// TIA Portal V20 export
// export: Created 2026-10-20T18:54:16.3544517Z, ExportSetting None, DisplayName Totally Integrated Automation Portal, DisplayVersion V20 Update 6, DisplayName TIA Portal Openness, DisplayVersion V20 Update 6, DisplayName TIA Portal Version Control Interface, DisplayVersion V20 Update 6, DisplayName SINAMICS Startdrive Advanced, DisplayVersion V20 SP1, DisplayName SINAMICS Startdrive G130, G150, S120, S150, SINAMICS MV, G220, S200, S210, DisplayVersion V20 SP1, DisplayName SINAMICS Startdrive G110M, G120, G120C, G120D, G120P, G115D, DisplayVersion V20 SP1, DisplayName STEP 7 Professional, DisplayVersion V20 Update 6, DisplayName STEP 7 Safety, DisplayVersion V20 Update 2, DisplayName WinCC Basic/Comfort/Advanced, DisplayVersion V20 Update 6, DisplayName WinCC Unified, DisplayVersion V20 Update 6
VAR_GLOBAL   // PLC tag table "IO_Main Panel"
   "MAIN PANEL STACK LIGHT RED" AT %Q350.0 : Bool;   // TESTED
   "MAIN PANEL STACK LIGHT AMBER" AT %Q350.1 : Bool;   // TESTED
   "MAIN PANEL STACK LIGHT GREEN" AT %Q350.2 : Bool;   // TESTED
   "SCA 1002 REMOTE PANEL SUPPLY FEEDBACK" AT %I300.0 : Bool;   // TESTED
   "SCA 2002 REMOTE PANEL SUPPLY FEEDBACK" AT %I300.1 : Bool;
   "SCA 3002 REMOTE PANEL SUPPLY FEEDBACK" AT %I300.2 : Bool;
   "SCA 4001 REMOTE PANEL SUPPLY FEEDBACK" AT %I300.3 : Bool;
   "SCA 5001 REMOTE PANEL SUPPLY FEEDBACK" AT %I300.4 : Bool;
   "SW1 SWITCH PANEL SUPPLY FEEDBACK" AT %I300.5 : Bool;
   "SW2 SWITCH PANEL SUPPLY FEEDBACK" AT %I300.6 : Bool;
   "SW3 SWITCH PANEL SUPPLY FEEDBACK" AT %I300.7 : Bool;
   "60TA1 PSU 24V OK FEEDBACK" AT %I301.0 : Bool;   // IT WILL NEVER GO TO FALSE
   "60TA2 PSU 24V OK FEEDBACK" AT %I301.1 : Bool;   // IT WILL NEVER GO TO FALSE
   "441FC1 CHARGER PANEL 1 SUPPLY FEEDBACK" AT %I301.2 : Bool;
   "441FC2 CHARGER PANEL 2 SUPPLY FEEDBACK" AT %I301.3 : Bool;
   "441FC3 CHARGER PANEL 3 SUPPLY FEEDBACK" AT %I301.4 : Bool;
   "41FC1 COOLING FAN MCB FEEDBACK" AT %I301.5 : Bool;   // TESTED
   "62TA1 PSU 48V OK FEEDBACK" AT %I301.6 : Bool;   // TESTED
   "CHARGER PANELS 4,5,6,7,8 SUPPLY FEEDBACK" AT %I301.7 : Bool;   // 441FC4, 442FC1, 442FC2, 442FC3, 442FC4
   "EMERGENCY STOP (CABINET) - CH1" AT %I320.0 : Bool;   // TESTED
   "EMERGENCY STOP RESET (CABINET)" AT %I320.1 : Bool;   // TESTED
   "EMERGENCY STOP (CABINET) - CH2" AT %I321.0 : Bool;   // TESTED
   "RESET PLC HMI - CH2" AT %Q350.4 : Bool;
   "RESET PLC HMI - CH1" AT %Q350.3 : Bool;
   "PLC_HMI - Profinet_Error_HMI 1" AT %I330.6 : Bool;
   "PLC_HMI - Profinet_Error_HMI 2" AT %I330.7 : Bool;
   "PLC_HMI - HMI 2 Estop" AT %I329.7 : Bool;
   "PLC_HMI - HMI 1 Estop" AT %I329.6 : Bool;
END_VAR
